(* IEC 61131-3 sources: model-first-plc-agent-ai/results/T4-W-22, 2 files *)

(* ---- a1_code.st ---- *)
FUNCTION_BLOCK LevelControlRuntime
VAR_INPUT
    StartSignal : BOOL;
    StopSignal : BOOL;
    LevelSample : INT;
    FullScaleValue : INT;
    h_span : REAL;
    Kp : REAL;
    Ti : REAL;
    Td : REAL;
    t_h : TIME;
    CycleSeconds : REAL;
END_VAR
VAR_OUTPUT
    FillCommand : INT;
    DischargeCommand : INT;
    fill_valve : BOOL;
    discharge_valve : BOOL;
END_VAR
VAR CONSTANT
    REGION_LOW : INT := 0;
    REGION_MIDDLE : INT := 1;
    REGION_HIGH : INT := 2;
END_VAR
VAR
    StartEdge : R_TRIG;
    HoldTimer : TON;

    start : BOOL;
    stop : BOOL;
    settled : BOOL;
    r : INT := 0;

    x0 : BOOL := TRUE;
    x1 : BOOL := FALSE;
    WasRegulating : BOOL;

    h : REAL;
    h_sp : REAL;
    h_target : REAL;
    h_max : REAL;
    eps : REAL;
    LevelError : REAL;
    PreviousError : REAL := 0.0;

    ProportionalTerm : REAL;
    IntegralTerm : REAL := 0.0;
    DerivativeTerm : REAL;
    CandidateIntegral : REAL;
    UnconstrainedDemand : REAL;
    CandidateDemand : REAL;
    LimitedDemand : REAL;
END_VAR

StartEdge(CLK := StartSignal);
start := StartEdge.Q;
stop := StopSignal;

h_sp := 0.8 * h_span;
h_target := h_sp;
h_max := 0.9 * h_span;
eps := 0.02 * h_span;

h := INT_TO_REAL(LevelSample) * h_span / INT_TO_REAL(FullScaleValue);
LevelError := h_sp - h;

IF h < h_target THEN
    r := REGION_LOW;
ELSIF h < h_max THEN
    r := REGION_MIDDLE;
ELSE
    r := REGION_HIGH;
END_IF;

WasRegulating := x1;

(* The hold condition measures continuous time inside the tolerance
   band while x1 is active, not merely the duration of x1. *)
HoldTimer(
    IN := x1 AND NOT stop AND (ABS(LevelError) <= eps),
    PT := t_h
);
settled := HoldTimer.Q;

(* Evaluate transitions using the situation at the start of this scan. *)
IF x0 THEN
    IF start AND NOT stop AND NOT (r = REGION_HIGH) THEN
        x0 := FALSE;
        x1 := TRUE;
    END_IF;
ELSIF x1 THEN
    IF stop OR settled OR (r = REGION_HIGH) THEN
        x1 := FALSE;
        x0 := TRUE;
    END_IF;
END_IF;

(* Clear the owned hold condition immediately upon leaving x1. *)
IF NOT x1 THEN
    HoldTimer(IN := FALSE, PT := t_h);
    settled := FALSE;
END_IF;

fill_valve := x1;
discharge_valve := x1;

FillCommand := 0;
DischargeCommand := 0;
LimitedDemand := 0.0;

(* PID demand is expressed as a fraction of full valve opening.
   Kp therefore has units of opening fraction per level unit.
   Ti, Td, and CycleSeconds are expressed in seconds. *)
IF x1 THEN
    IF NOT WasRegulating THEN
        PreviousError := LevelError;
    END_IF;

    ProportionalTerm := Kp * LevelError;
    DerivativeTerm := 0.0;

    IF (Td > 0.0) AND (CycleSeconds > 0.0) THEN
        DerivativeTerm :=
            Kp * Td * (LevelError - PreviousError) / CycleSeconds;
    END_IF;

    UnconstrainedDemand :=
        ProportionalTerm + IntegralTerm + DerivativeTerm;

    (* Suspend integration whenever the current output is clamped.
       Also reject an integral update that would cause clamping. *)
    IF (Ti > 0.0) AND (CycleSeconds > 0.0) THEN
        IF (UnconstrainedDemand >= 0.0) AND
           (UnconstrainedDemand <= 1.0) THEN
            CandidateIntegral :=
                IntegralTerm + Kp * LevelError * CycleSeconds / Ti;
            CandidateDemand :=
                ProportionalTerm + CandidateIntegral + DerivativeTerm;

            IF (CandidateDemand >= 0.0) AND
               (CandidateDemand <= 1.0) THEN
                IntegralTerm := CandidateIntegral;
            END_IF;
        END_IF;
    END_IF;

    UnconstrainedDemand :=
        ProportionalTerm + IntegralTerm + DerivativeTerm;

    IF UnconstrainedDemand < 0.0 THEN
        LimitedDemand := 0.0;
    ELSIF UnconstrainedDemand > 1.0 THEN
        LimitedDemand := 1.0;
    ELSE
        LimitedDemand := UnconstrainedDemand;
    END_IF;

    FillCommand :=
        REAL_TO_INT(LimitedDemand * INT_TO_REAL(FullScaleValue));
    DischargeCommand :=
        REAL_TO_INT(0.4 * INT_TO_REAL(FullScaleValue));
END_IF;

(* IntegralTerm is retained, but never integrated, outside x1. *)
PreviousError := LevelError;

END_FUNCTION_BLOCK

PROGRAM Main
VAR
    StartCommand AT %IX100.0 : BOOL;
    StopCommand AT %IX100.1 : BOOL;
    LevelMeter AT %IW100 : INT;
    FillValve AT %QW100 : INT;
    DischargeValve AT %QW101 : INT;
END_VAR
VAR CONSTANT
    FULL_SCALE : INT := 1000;
    ScanSeconds : REAL := 0.02;
END_VAR
VAR
    Controller : LevelControlRuntime;

    h_span : REAL := 10.0;
    t_h : TIME := T#10s;

    (* Initial tuning values; commission for the simulated plant. *)
    Kp : REAL := 1.0;
    Ti : REAL := 10.0;
    Td : REAL := 0.0;
END_VAR

Controller(
    StartSignal := StartCommand,
    StopSignal := StopCommand,
    LevelSample := LevelMeter,
    FullScaleValue := FULL_SCALE,
    h_span := h_span,
    Kp := Kp,
    Ti := Ti,
    Td := Td,
    t_h := t_h,
    CycleSeconds := ScanSeconds
);

FillValve := Controller.FillCommand;
DischargeValve := Controller.DischargeCommand;

END_PROGRAM

CONFIGURATION Config0
    RESOURCE Res0 ON PLC
        TASK ControlTask(INTERVAL := T#20ms, PRIORITY := 0);
        PROGRAM MainInstance WITH ControlTask : Main;
    END_RESOURCE
END_CONFIGURATION

(* ---- a2_code.st ---- *)
FUNCTION_BLOCK FB_LevelControl
VAR_INPUT
    StartCommand : BOOL;
    StopCommand : BOOL;
    LevelMeter : INT;
    Kp : REAL;
    Ti : REAL;
    Td : REAL;
    cycle_seconds : REAL;
END_VAR
VAR_OUTPUT
    FillValve : INT;
    DischargeValve : INT;
    fill_valve : BOOL;
    discharge_valve : BOOL;
END_VAR
VAR CONSTANT
    FULL_SCALE : INT := 1000;
    h_span : REAL := 10.0;
    h_sp : REAL := 8.0;
    h_target : REAL := 8.0;
    h_max : REAL := 9.0;
    eps : REAL := 0.2;
    t_h : TIME := T#10s;
    REGION_LOW : INT := 0;
    REGION_MIDDLE : INT := 1;
    REGION_HIGH : INT := 2;
END_VAR
VAR
    start_edge : R_TRIG;
    hold_timer : TON;
    start : BOOL;
    stop : BOOL;
    settled : BOOL;
    r : INT;
    active_state : INT := 0;
    was_regulating : BOOL := FALSE;
    h : REAL;
    error_value : REAL;
    previous_error : REAL := 0.0;
    integral_value : REAL := 0.0;
    candidate_integral : REAL;
    derivative_value : REAL;
    raw_demand : REAL;
    limited_demand : REAL;
END_VAR

start_edge(CLK := StartCommand);
start := start_edge.Q;
stop := StopCommand;

h := INT_TO_REAL(LevelMeter) * h_span / INT_TO_REAL(FULL_SCALE);
error_value := h_sp - h;

IF h < h_target THEN
    r := REGION_LOW;
ELSIF h < h_max THEN
    r := REGION_MIDDLE;
ELSE
    r := REGION_HIGH;
END_IF;

hold_timer(
    IN := (active_state = 1) AND NOT stop
          AND (ABS(error_value) <= eps),
    PT := t_h
);
settled := hold_timer.Q;

IF stop THEN
    active_state := 0;
ELSE
    CASE active_state OF
        0:
            IF start THEN
                active_state := 1;
            END_IF;
        1:
            IF settled OR (r = REGION_HIGH) THEN
                active_state := 0;
            END_IF;
    ELSE
        active_state := 0;
    END_CASE;
END_IF;

(* Apply the overfill termination immediately, including on entry. *)
IF (active_state = 1) AND (r = REGION_HIGH) THEN
    active_state := 0;
END_IF;

fill_valve := (active_state = 1);
discharge_valve := (active_state = 1);

FillValve := 0;
DischargeValve := 0;

IF fill_valve THEN
    IF NOT was_regulating THEN
        integral_value := 0.0;
        previous_error := error_value;
    END_IF;

    derivative_value := 0.0;
    IF cycle_seconds > 0.0 THEN
        derivative_value :=
            Kp * Td * (error_value - previous_error) / cycle_seconds;
    END_IF;

    (* PID demand uses a normalized opening: 0.0 through 1.0. *)
    candidate_integral := integral_value;
    IF (Ti > 0.0) AND (cycle_seconds > 0.0) THEN
        candidate_integral :=
            integral_value + Kp * error_value * cycle_seconds / Ti;
    END_IF;

    raw_demand :=
        Kp * error_value + candidate_integral + derivative_value;

    (* Do not commit the integral update when the demand is clamped. *)
    IF raw_demand > 1.0 THEN
        limited_demand := 1.0;
    ELSIF raw_demand < 0.0 THEN
        limited_demand := 0.0;
    ELSE
        limited_demand := raw_demand;
        integral_value := candidate_integral;
    END_IF;

    previous_error := error_value;
    FillValve :=
        REAL_TO_INT(limited_demand * INT_TO_REAL(FULL_SCALE));
    DischargeValve :=
        REAL_TO_INT(0.4 * INT_TO_REAL(FULL_SCALE));
ELSE
    integral_value := 0.0;
    previous_error := error_value;
END_IF;

was_regulating := fill_valve;

END_FUNCTION_BLOCK

PROGRAM Main
VAR
    StartCommand AT %IX100.0 : BOOL;
    StopCommand AT %IX100.1 : BOOL;
    LevelMeter AT %IW100 : INT;
    FillValve AT %QW100 : INT;
    DischargeValve AT %QW101 : INT;
END_VAR
VAR
    controller : FB_LevelControl;
    (* Commission these gains for the simulated plant. *)
    Kp : REAL := 1.0;
    Ti : REAL := 5.0;
    Td : REAL := 0.0;
    cycle_seconds : REAL := 0.02;
    fill_valve : BOOL;
    discharge_valve : BOOL;
END_VAR

controller(
    StartCommand := StartCommand,
    StopCommand := StopCommand,
    LevelMeter := LevelMeter,
    Kp := Kp,
    Ti := Ti,
    Td := Td,
    cycle_seconds := cycle_seconds
);

FillValve := controller.FillValve;
DischargeValve := controller.DischargeValve;
fill_valve := controller.fill_valve;
discharge_valve := controller.discharge_valve;

END_PROGRAM

CONFIGURATION Config0
    RESOURCE Res0 ON PLC
        TASK MainTask(INTERVAL := T#20ms, PRIORITY := 0);
        PROGRAM MainInstance WITH MainTask : Main;
    END_RESOURCE
END_CONFIGURATION
